SUBAPPLICATION PAGE (* Subapplication Type *)
  (* Standard: 61499-2 *)
  (* Version 1.0, 2023-02-07, franz *)
  IMPORT isobus::UT::io::Auxiliary::IN::AuxiliaryState::AuxDisabled;
  IMPORT isobus::UT::io::Button::ButtonActivationCode::BT_RELEASED_UNLATCHED;
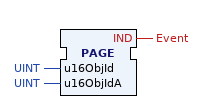
  EVENT_OUTPUT
    IND;
  END_EVENT
  VAR_INPUT
    u16ObjId : UINT;
    u16ObjIdA : UINT;
  END_VAR
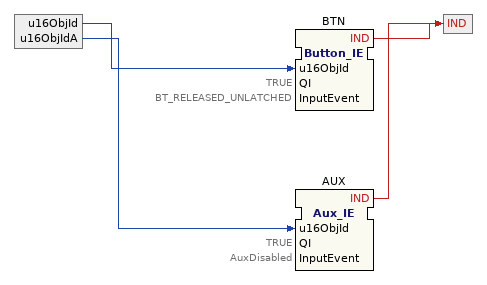
  FBS
    BTN : isobus::UT::io::Button::Button_IE(QI := TRUE, InputEvent := BT_RELEASED_UNLATCHED);
    AUX : isobus::UT::io::Auxiliary::IN::Aux_IE(QI := TRUE, InputEvent := AuxDisabled);
  END_FBS
  EVENT_CONNECTIONS
    AUX.IND TO IND;
    BTN.IND TO IND;
  END_CONNECTIONS
  DATA_CONNECTIONS
    u16ObjId TO BTN.u16ObjId;
    u16ObjIdA TO AUX.u16ObjId;
  END_CONNECTIONS
END_SUBAPPLICATION
